// TIA Portal V20 export
// export: Created 2026-10-20T12:46:26.647728Z, ExportSetting WithDefaults, DisplayName Totally Integrated Automation Portal, DisplayVersion V20 Update 6, DisplayName TIA Portal Openness, DisplayVersion V20 Update 6, DisplayName TIA Portal Version Control Interface, DisplayVersion V20 Update 6, DisplayName SINAMICS Startdrive Advanced, DisplayVersion V20 SP1, DisplayName SINAMICS Startdrive G130, G150, S120, S150, SINAMICS MV, G220, S200, S210, DisplayVersion V20 SP1, DisplayName SINAMICS Startdrive G110M, G120, G120C, G120D, G120P, G115D, DisplayVersion V20 SP1, DisplayName STEP 7 Professional, DisplayVersion V20 Update 6, DisplayName STEP 7 Safety, DisplayVersion V20 Update 2, DisplayName WinCC Basic/Comfort/Advanced, DisplayVersion V20 Update 6, DisplayName WinCC Unified, DisplayVersion V20 Update 6
DATA_BLOCK "CNV_HMI"   // DB40
{ S7_Optimized_Access := 'TRUE' }
VERSION : 0.1
// stored: AutoNumber true, DBAccessibleFromOPCUA true, IsOnlyStoredInLoadMemory false, IsRetainMemResEnabled false, IsWriteProtectedInAS false, MemoryReserve 100
   VAR
      "Manual_Sfty_Stopper_Up(1)" : Array[1..5] of Bool;
      "Manual_Sfty_Stopper_Down(1)" : Array[1..5] of Bool;
      In_Out : Array[1..5] of Bool;
      ID : Array[1..5] of DInt;
      "Task_ID(1)" : Array[1..5] of UInt;
      Manual_Bwd : Array[1..5] of Bool;
      "Reset(1)" : Array[1..5] of Bool;
      "Pallet_Type(1)" : Array[1..5] of UInt;
      Manual_Fwd : Array[1..5] of Bool;
      Enable : Array[1..5] of Bool;
      "Pallet_Align_Right(1)" : Array[1..5] of Bool;
      "Enable(1)" : Array[1..5] of Bool;
      Pallet_Type : Array[1..5] of UInt;
      Pallet_Allignment : Array[1..5] of Bool;
      "Transfer_To_ID(1)" : Array[1..5] of DInt;
      Pallet_Align_Right : Array[1..5] of Bool;
      "Manual_Bwd(1)" : Array[1..5] of Bool;
      "Pallet_Align_Left(1)" : Array[1..5] of Bool;
      Reset : Array[1..5] of Bool;
      Stop : Array[1..5] of Bool;
      Pallet_Align_Center : Array[1..5] of Bool;
      "Stop(1)" : Array[1..5] of Bool;
      "Start_Transfer(1)" : Array[1..5] of Bool;
      Pallet_Align_Left : Array[1..5] of Bool;
      Start_Transfer : Array[1..5] of Bool;
      "ID(1)" : Array[1..5] of DInt;
      "Transfer_From_ID(1)" : Array[1..5] of DInt;
      "Manual_Fwd(1)" : Array[1..5] of Bool;
      Mode_Change : Array[1..5] of UInt;
      Transfer_To_ID : Array[1..5] of DInt;
      "Mode_Change(1)" : Array[1..5] of UInt;
      Transfer_From_ID : Array[1..5] of DInt;
      UpDown : Array[1..5] of UInt;
      Same_Cnv : Array[1..5] of Bool;
      CNV2_Selected : Array[1..5] of UInt;
      "Pallet_Allignment(1)" : Array[1..5] of Bool;
      "Occupied(1)" : Array[1..5] of Bool;
      Mode : Array[1..5] of UInt;
      "Running(1)" : Array[1..5] of Bool;
      "Enabled(1)" : Array[1..5] of Bool;
      Motor_Speed_Actual : Array[1..5] of UInt;
      Running : Array[1..5] of Bool;
      "SM_State(1)" : Array[1..5] of UInt;
      "Warning(1)" : Array[1..5] of UInt;
      Stopped : Array[1..5] of Bool;
      Enabled : Array[1..5] of Bool;
      Error : Array[1..5] of Bool;
      "Motor_Speed_Requested(1)" : Array[1..5] of UInt;
      Current_Task_ID : Array[1..5] of UInt;
      "Mode(1)" : Array[1..5] of UInt;
      "Current_Task_Type(1)" : Array[1..5] of UInt;
      Warning : Array[1..5] of UInt;
      "Current_Task_ID(1)" : Array[1..5] of UInt;
      Current_Task_Type : Array[1..5] of UInt;
      "Stopped(1)" : Array[1..5] of Bool;
      Motor_Direction : Array[1..5] of UInt;
      SM_State : Array[1..5] of UInt;
      "Ready_For_Task(1)" : Array[1..5] of Bool;
      Ready_For_Task : Array[1..5] of Bool;
      Occupied : Array[1..5] of Bool;
      "Error(1)" : Array[1..5] of Bool;
      Shuttle_in_place : Array[1..5] of Bool;
      Motor_Speed_Requested : Array[1..5] of UInt;
      "Motor_Direction(1)" : Array[1..5] of UInt;
      "Motor_Speed_Actual(1)" : Array[1..5] of UInt;
      "Shuttle_in_place(1)" : Array[1..5] of Bool;
      Motor_Ready : Array[1..5] of Bool;
      "Motor_Current_Actual(1)" : Array[1..5] of Real;
      Motor_Status : Array[1..5] of UInt;
      "Motor_Status(1)" : Array[1..5] of UInt;
      Motor_Current_Actual : Array[1..5] of Real;
      "Motor_Ready(1)" : Array[1..5] of Bool;
      Task_ID : Array[1..5] of UInt;
      Level_Selected : Array[1..5] of UInt;
      "UpDown(1)" : Array[1..5] of UInt;
      Motor_Actual_Torque : Array[1..5] of Real;
      "Motor_Actual_Torque(1)" : Array[1..5] of Real;
      Safety_OK : Array[1..5] of Bool;
      Reset_Comissioning : Array[1..5] of Bool;
      Charge_Commands : Array[1..5] of Bool;
      Charge_Cnv : Array[1..5] of Bool;
      Reset_All : Array[1..5] of Bool;
      Sdetect1 : Array[1..5] of Bool;
      Sdetect2 : Array[1..5] of Bool;
      "Sdetect1(1)" : Array[1..5] of Bool;
      "Sdetect2(1)" : Array[1..5] of Bool;
      "Rpd2(1)" : Array[1..5] of Bool;
      Center : Array[1..5] of Bool;
      "Rpd1(1)" : Array[1..5] of Bool;
      "Lpd2(1)" : Array[1..5] of Bool;
      "Lpd1(1)" : Array[1..5] of Bool;
      Rpd1 : Array[1..5] of Bool;
      Lpd1 : Array[1..5] of Bool;
      Rpd2 : Array[1..5] of Bool;
      "Right(1)" : Array[1..5] of Bool;
      Right : Array[1..5] of Bool;
      Left : Array[1..5] of Bool;
      "Left(1)" : Array[1..5] of Bool;
   END_VAR
BEGIN
END_DATA_BLOCK
